{attribute 'qualified_only'}
{attribute 'strict'}
{attribute 'to_string'}
TYPE E_HttpExporterState :
(
	error := -10,
	idle := 0,
	serializing := 10,
	sending := 20,
	waiting := 30,
	processing := 40,
	done := 99
);
END_TYPE
//  error = '-10'

(* stored: Version 1.1.0.1
   EnumerationTextList E_HttpExporterState: Id {35159dc4-d259-4d27-9ff6-b0fff5699231} *)
